Yaskawa INFORM job: DROPPAR.JBI

/JOB
//NAME DROPPAR
//POS
///NPOS 4,0,0,0,0,0
///TOOL 9
///POSTYPE PULSE
///PULSE
C00000=-56,2,2,0,0,0
C00001=-104,-5,-32,29,30,64
///TOOL 9
///POSTYPE BASE
///RECTAN
///RCONF 0,0,0,1,0,0,0,0
C00002=-345.000,-1635.000,230.000,90.00,-0.00,0.00
C00003=-345.000,-1175.000,480.000,90.00,-0.00,0.00
//INST
///DATE 2026/10/26 01:19
///COMM Generated using RoboDK
///ATTR SC,RW,RJ
///GROUP1 RB1
NOP
'Using Table (targets wrt base
'):
'0.0,-1500.0,-60.0,0.0,0.0,0.0
'Setting Tool 9 (Wood_Holder):
SETE P00095 (1) 0
SETE P00095 (2) 0
SETE P00095 (3) 40000
SETE P00095 (4) 0
SETE P00095 (5) 0
SETE P00095 (6) 0
SETTOOL TL#(9) P00095
MOVJ C00000 VJ=50.00
MOVJ C00001 VJ=50.00
MOVL C00002 V=1000.0
'Detach from Wood_Holder
'Detach from Wood_Holder
MOVL C00003 V=1000.0
END
